// TIA Portal V21 export
// export: Created 2026-11-11T00:48:06.6609566Z, ExportSetting WithDefaults, DisplayName Totally Integrated Automation Portal, DisplayVersion V21 Update 3, DisplayName STEP 7 Professional, DisplayVersion V21 Update 3, DisplayName STEP 7 Safety, DisplayVersion V21, DisplayName Tech WebApplication, DisplayVersion V21, DisplayName WinCC Basic/Comfort/Advanced, DisplayVersion V21 Update 3, DisplayName WinCC Unified, DisplayVersion V21 Update 3
FUNCTION_BLOCK "FB_Scl_m107"   // FB297, SCL
{ S7_Optimized_Access := 'TRUE' }
VERSION : 0.1
// stored: AutoNumber true, IsIECCheckEnabled false, IsRetainMemResEnabled false, MemoryReserve 100, SetENOAutomatically false, UDAEnableTagReadback false
   VAR_INPUT
      vin : Variant;
      dba : DB_ANY;
   END_VAR
   VAR_IN_OUT
      by8 : Array[0..99] of Byte;
      arrA : Array[0..9] of Int;
      arrB : Array[0..9] of Int;
      barr : Array[0..15] of Bool;
      va : Array[*] of Int;
      pos : DInt;
   END_VAR
   VAR
      t1 { S7_SetPoint := 'True'} : TON_TIME;
      mem : LReal;
   END_VAR
   VAR_TEMP
      i : Int;
      di : DInt;
      r : Real;
      lr : LReal;
      w : Word;
      dw : DWord;
      "b" : Bool;
      "by" : Byte;
      t : Time;
      ec : Int;
      o0 : Int;
      o1 : Int;
      v : Variant;
   END_VAR
BEGIN
   DEMUX(K := #di, IN := #i, OUT0 => #o0, OUT1 => #o1);
END_FUNCTION_BLOCK
